// Generated by voz_llm_plc_agent
// Target: Siemens TIA Portal V18 - SCL external source
// Review and compile before any download to physical hardware.

FUNCTION_BLOCK "PLC_PRG"
{ S7_Optimized_Access := 'TRUE' }
VERSION : 0.1
VAR_INPUT
   I_Mode_Manual : Bool := FALSE;
   I_Manual_Motor_Command : Bool := FALSE;
   I_Automatic_Motor_Command : Bool := FALSE;
   I_Emergency : Bool := FALSE;
END_VAR
VAR_OUTPUT
   Q_Motor_Enable : Bool := FALSE;
END_VAR
BEGIN
(* Salidas: contribucion automatica (secuencia/condiciones) y manual, con sus bloqueos *)
#Q_Motor_Enable := ((#I_Mode_Manual AND #I_Manual_Motor_Command) OR (NOT #I_Mode_Manual AND #I_Automatic_Motor_Command)) AND NOT FALSE;
(* Bloqueo: #I_Emergency fuerza a FALSE #Q_Motor_Enable de inmediato *)
IF #I_Emergency THEN
    #Q_Motor_Enable := FALSE;
END_IF;
END_FUNCTION_BLOCK

DATA_BLOCK "DB_PLC_PRG"
{ S7_Optimized_Access := 'TRUE' }
VERSION : 0.1
NON_RETAIN
"PLC_PRG"
BEGIN
END_DATA_BLOCK

ORGANIZATION_BLOCK "Main"
{ S7_Optimized_Access := 'TRUE' }
VERSION : 0.1
BEGIN
   "DB_PLC_PRG"(
      I_Mode_Manual := "I_Mode_Manual",
      I_Manual_Motor_Command := "I_Manual_Motor_Command",
      Q_Motor_Enable => "Q_Motor_Enable",
      I_Automatic_Motor_Command := "I_Automatic_Motor_Command",
      I_Emergency := "I_Emergency"
   );
END_ORGANIZATION_BLOCK
